(* IEC 61131-3 sources: kns-port-domestic/targets/astra/lib/src/DUTs/ControlValve, 5 files *)

(* ---- E_CvAlarm.dut.st ---- *)
// Назначение: индексы слотов тревог регулирующего клапана. Нестрогое перечисление: им
//             индексируются массивы.
// Автор:      kr0nsch
// Версия:     0.1.0
// Документ:   docs/fb/FB_ControlValve.md
{attribute 'qualified_only'}
TYPE E_CvAlarm :
(
    Deviation       := 0,   // рассогласование задания и ОС положения
    FbFailure       := 1,   // ОС положения недостоверна
    PositionerFault := 2,   // авария позиционера или канала AO
    InterlockAct    := 3    // действует блокировка (по умолчанию выключена)
) UINT;
END_TYPE

(* ---- E_CvFaultAction.dut.st ---- *)
// Назначение: реакция регулирующего клапана на отказ.
// Автор:      kr0nsch
// Версия:     0.1.0
// Документ:   docs/fb/FB_ControlValve.md
{attribute 'qualified_only'}
{attribute 'strict'}
TYPE E_CvFaultAction :
(
    Hold    := 0,   // удерживать положение
    SafePos := 1    // в rSafePos_pct без рампы
) INT;
END_TYPE

(* ---- ST_ControlValveCfg.dut.st ---- *)
// Назначение: параметры регулирующего клапана (Persistent Variables приложения,
//             VAR_IN_OUT CONSTANT stCfg). Значения по умолчанию проходят CheckConfig.
//             Тип лежит в Persistent Variables приложения и заморожен в пределах 1.x (A-13).
// Автор:      kr0nsch
// Версия:     0.1.0
// Документ:   docs/fb/FB_ControlValve.md
{attribute 'qualified_only'}
TYPE ST_ControlValveCfg :
STRUCT
    rOutMin_pct     : REAL := 0.0;     // нижний предел задания, %
    rOutMax_pct     : REAL := 100.0;   // верхний предел задания, %
    rRateUp_pctps   : REAL := 0.0;     // %/с; 0 — без ограничения
    rRateDown_pctps : REAL := 0.0;     // %/с; 0 — без ограничения
    rTightShut_pct  : REAL := 0.0;     // выход ниже порога → 0 % (плотное закрытие); 0 — выключено
    xOutInvert      : BOOL := FALSE;   // TRUE: 100 % хода = 4 мА
    rSafePos_pct    : REAL := 0.0;     // положение по блокировке и отказу (не путать с механическим)
    eFaultAction    : E_CvFaultAction := E_CvFaultAction.Hold;
    xFbUsed         : BOOL := FALSE;   // ОС положения подключена
    rDevMax_pct     : REAL := 5.0;     // допуск рассогласования, %
    tDev            : TIME := T#30S;   // задержка рассогласования
    xDevIsFault     : BOOL := FALSE;   // FALSE — рассогласование только предупреждение
    wInterlockMask  : WORD := 16#FFFF; // какие биты wInterlock действуют
    udiAlarmIdBase  : UDINT := 0;      // номер первой тревоги устройства (dev_no * 10)
    astAlarm        : ARRAY[0..GVL_Const.DEV_ALARMS_MAX - 1] OF ST_AlarmCfg := [
        (ePriority := E_AlarmPriority.Low),       // 0 Deviation
        (ePriority := E_AlarmPriority.Low),       // 1 FbFailure
        (ePriority := E_AlarmPriority.Medium),    // 2 PositionerFault
        (ePriority := E_AlarmPriority.None),      // 3 InterlockAct
        (ePriority := E_AlarmPriority.None), (ePriority := E_AlarmPriority.None),
        (ePriority := E_AlarmPriority.None), (ePriority := E_AlarmPriority.None)];
END_STRUCT
END_TYPE

(* ---- ST_ControlValveCmd.dut.st ---- *)
// Назначение: команды HMI/SCADA регулирующего клапана (GVL_Hmi приложения, VAR_IN_OUT stCmd).
// Автор:      kr0nsch
// Версия:     0.1.0
// Документ:   docs/fb/FB_ControlValve.md
{attribute 'qualified_only'}
TYPE ST_ControlValveCmd :
STRUCT
    stCommon      : ST_DeviceCmd;
    rPosSpMan_pct : REAL;   // задание в Manual, %; в Auto/Local/OOS ФБ пишет сюда текущий rOut_pct
END_STRUCT
END_TYPE

(* ---- ST_ControlValveSts.dut.st ---- *)
// Назначение: состояние регулирующего клапана для HMI/SCADA. 52 байта, 26 регистров Modbus:
//             только 16- и 32-битные поля без скрытого выравнивания.
// Автор:      kr0nsch
// Версия:     0.1.0
// Документ:   docs/fb/FB_ControlValve.md
{attribute 'qualified_only'}
TYPE ST_ControlValveSts :
STRUCT
    stCommon       : ST_DeviceSts;   // 0..27
    rPosSp_pct     : REAL;   // 28: задание после пределов, до рампы
    rOut_pct       : REAL;   // 32: задание положения, % хода
    rOut_mA        : REAL;   // 36: на AO с учётом инверсии
    rPosFb_pct     : REAL;   // 40: ОС положения
    rDeviation_pct : REAL;   // 44: rOut_pct − rPosFb_pct
    wInterlock     : WORD;   // 48: действующие блокировки
    uiFirstOut     : UINT;   // 50: первопричина блокировки; NO_FIRST_OUT — нет
END_STRUCT
END_TYPE
